// Tests for HalfBROT.F_FocusTrackStoredPosition (HalfBROT 0.7.2, #66): when the stored focus position takes the actual position.
FUNCTION_BLOCK F_FocusTrackStoredPosition_Tests EXTENDS TcUnit.FB_TestSuite
VAR
END_VAR

Calibrated_Locked_Idle_Tracks();
Unlocked_Does_Not_Track();
Homing_Does_Not_Track();
Not_Calibrated_Does_Not_Track();

// #66: the function has no mode input. A focus jogged in manual mode is stored like one moved in automatic mode.
METHOD PRIVATE Calibrated_Locked_Idle_Tracks
VAR
END_VAR
TEST('Calibrated_Locked_Idle_Tracks');
AssertTrue(Condition := HalfBROT.F_FocusTrackStoredPosition(bCalibrated := TRUE, bLocked := TRUE, bHoming := FALSE), Message := 'calibrated, locked, not homing');
TEST_FINISHED();
END_METHOD

// While the drive is enabled the focus moves or is about to.
METHOD PRIVATE Unlocked_Does_Not_Track
VAR
END_VAR
TEST('Unlocked_Does_Not_Track');
AssertFalse(Condition := HalfBROT.F_FocusTrackStoredPosition(bCalibrated := TRUE, bLocked := FALSE, bHoming := FALSE), Message := 'unlocked');
TEST_FINISHED();
END_METHOD

// The homing owns fLastPosition (MC_Direct reads it).
METHOD PRIVATE Homing_Does_Not_Track
VAR
END_VAR
TEST('Homing_Does_Not_Track');
AssertFalse(Condition := HalfBROT.F_FocusTrackStoredPosition(bCalibrated := TRUE, bLocked := TRUE, bHoming := TRUE), Message := 'homing');
TEST_FINISHED();
END_METHOD

// An uncalibrated focus has no valid actual position.
METHOD PRIVATE Not_Calibrated_Does_Not_Track
VAR
END_VAR
TEST('Not_Calibrated_Does_Not_Track');
AssertFalse(Condition := HalfBROT.F_FocusTrackStoredPosition(bCalibrated := FALSE, bLocked := TRUE, bHoming := FALSE), Message := 'not calibrated');
TEST_FINISHED();
END_METHOD

END_FUNCTION_BLOCK

(* stored: Version 1.1.0.1, ProductVersion 3.1.4024.15
   POU F_FocusTrackStoredPosition_Tests: Id {7bd749d6-1509-476c-9de3-2a7826d3900f}, SpecialFunc None
   Method Calibrated_Locked_Idle_Tracks: Id {c234a005-5ad7-4cc6-88bb-9b738a644373}
   Method Unlocked_Does_Not_Track: Id {c18ed53f-9c6c-48e4-b15f-1833acc4d89b}
   Method Homing_Does_Not_Track: Id {91dd4f63-beae-408f-8678-e9e7f5bbe9ee}
   Method Not_Calibrated_Does_Not_Track: Id {3a45cd72-43d7-4ee5-9da7-41e1db6ffef0} *)
